// TIA Portal V19 export
// export: Created 2026-10-19T00:00:00.0000000Z, ExportSetting None
FUNCTION_BLOCK "FB_ProbeLd"   // FB1, LAD
TITLE = FB_ProbeLd
{ S7_Optimized_Access := 'TRUE' }
// LD FB_ProbeLd → LAD (c2s7)
// stored: AutoNumber true, MemoryReserve 100, SetENOAutomatically false
   VAR_INPUT
      xStart : Bool;
      xStop : Bool;
      xPermit : Bool;
      iSp : Int;
   END_VAR
   VAR_OUTPUT
      xRun : Bool;
      iOut : Int;
      xMoved : Bool;
      xRunInv : Bool;
   END_VAR
   VAR
      _c2s7_xStart_P : Bool;
      _c2s7_xStop_N : Bool;
   END_VAR
   VAR_TEMP
      _c2s7_xStart_e : Bool;
      _c2s7_xStop_e : Bool;
   END_VAR
   VAR_TEMP   // added for the SCL form of the ladder/FBD networks
      _w1 : Bool;
   END_VAR
BEGIN

REGION Network 1: Пуск по фронту
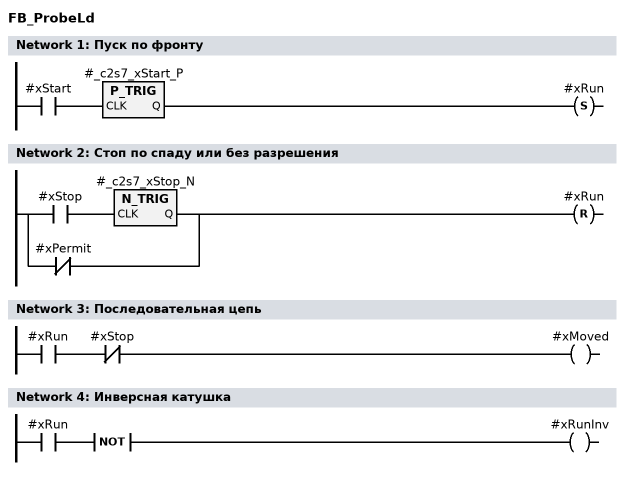
   RUNG wire#powerrail
      Contact( #xStart )
      P_Trig( #_c2s7_xStart_P )
      S_Coil( #xRun )
   END_RUNG
   // the same network as SCL:
   #_w1 := #xStart AND NOT #_c2s7_xStart_P;   // rising edge
   #_c2s7_xStart_P := #xStart;
   IF #_w1 THEN #xRun := TRUE; END_IF;
END_REGION

REGION Network 2: Стоп по спаду или без разрешения
   RUNG wire#powerrail
      Contact( #xStop )
      N_Trig( #_c2s7_xStop_N )
      wire#w1
      R_Coil( #xRun )
   END_RUNG
   RUNG wire#powerrail
      I_Contact( #xPermit )
   END_RUNG wire#w1
   // the same network as SCL:
   #_w1 := NOT #xStop AND #_c2s7_xStop_N;   // falling edge
   #_c2s7_xStop_N := #xStop;
   IF #_w1 OR NOT #xPermit THEN #xRun := FALSE; END_IF;
END_REGION

REGION Network 3: Последовательная цепь
   RUNG wire#powerrail
      Contact( #xRun )
      I_Contact( #xStop )
      Coil( #xMoved )
   END_RUNG
   // the same network as SCL:
   #xMoved := #xRun AND NOT #xStop;
END_REGION

REGION Network 4: Инверсная катушка
   RUNG wire#powerrail
      Contact( #xRun )
      Not()
      Coil( #xRunInv )
   END_RUNG
   // the same network as SCL:
   #xRunInv := NOT #xRun;
END_REGION
END_FUNCTION_BLOCK
